Fanuc KAREL source: kt00604.KL

-- PROVISIONAL review KL for V1013-1; original PC SHA256 7fb5911342036439b09a6b4d88e4647e6d12ce009c1241ad35af3e58da75da51
-- Incomplete behavior may be omitted. Consult companion uncertainty JSON. Do not deploy.
PROGRAM KT00604
%NOLOCKGROUP
VAR
  I1 : INTEGER
  I2 : INTEGER
  OUT : INTEGER
BEGIN
  -- UNRESOLVED_PC offsets 5-16; opcodes 2E,23
  -- UNRESOLVED_PC offsets 21-32; opcodes 2E,23
  -- UNRESOLVED_PC offsets 37-48; opcodes 2E,23
  -- UNRESOLVED_PC offsets 53-64; opcodes 2E,23
  -- UNRESOLVED_PC offsets 69-82; opcodes 21,51,23
  -- UNRESOLVED_PC offsets 87-91; opcodes 7F
END KT00604
